FUNCTION fShutterCmdSwitch  : stShutterCmdEvent
VAR_IN_OUT
	CmdEvent  : stShutterCmdEvent;
END_VAR
VAR_INPUT
	OpenSwitchState : stSwitchState;
    CloseSwitchState : stSwitchState;
    ShutterStateType : eShutterStateType;
END_VAR
VAR
END_VAR


// Exit if both switches are idle
IF OpenSwitchState.StateType = eSwitchStateType.IDLE AND
   CloseSwitchState.StateType = eSwitchStateType.IDLE THEN
    RETURN;
END_IF

// If shutter is moving and any switch was pressed
IF ShutterStateType <> eShutterStateType.IDLE THEN
    CmdEvent.Cmd.CmdType := eShutterCmdType.STOP;
// Double Open click
ELSIF (OpenSwitchState.StateType = eSwitchStateType.MULTI_CLICK) AND (OpenSwitchState.PressCount = 2) THEN
    CmdEvent.Cmd.CmdType := eShutterCmdType.OPEN;
// Double Close click
ELSIF (CloseSwitchState.StateType = eSwitchStateType.MULTI_CLICK) AND (CloseSwitchState.PressCount = 2) THEN
    CmdEvent.Cmd.CmdType := eShutterCmdType.CLOSE;
// Short Open click
ELSIF OpenSwitchState.StateType = eSwitchStateType.SHORT_CLICK THEN
    CmdEvent.Cmd.CmdType := eShutterCmdType.STEP_OPEN;
// Short Close click
ELSIF CloseSwitchState.StateType = eSwitchStateType.SHORT_CLICK THEN
    CmdEvent.Cmd.CmdType := eShutterCmdType.STEP_CLOSE;
// Long Open click
ELSIF OpenSwitchState.StateType = eSwitchStateType.LONG_CLICK THEN
    CmdEvent.Cmd.CmdType := eShutterCmdType.MOVE_TO_POSITION;
    CmdEvent.Cmd.Position := OpenLongClickPosition;
// Long Close click
ELSIF CloseSwitchState.StateType = eSwitchStateType.LONG_CLICK THEN
    CmdEvent.Cmd.CmdType := eShutterCmdType.MOVE_TO_POSITION;
    CmdEvent.Cmd.Position := CloseLongClickPosition;
END_IF

CmdEvent.Execute := TRUE;
CmdEvent.Source := eShutterCmdSource.SWITCH;

END_FUNCTION

(* stored: Version 1.1.0.1
   POU fShutterCmdSwitch: Id {69844d14-14f3-4a48-817d-2a200cd29af3}, SpecialFunc None *)
